// TIA Portal project "PLC_FB_Portfolio" (V14)

(* hardware
DEVICE "S71500/ET200MP station_1"  S7-1500 station
   slot 0: "Rail_0"  Rack  6ES7 590-1***0-0AA0
   slot 1: "PLC_1"  CPU 1511-1 PN  6ES7 511-1AK01-0AB0  V2.1
      slot 3: "CPU display_1"  6ES7591-1AA00-0AA0
*)

// ===== PLC "PLC_1"  CPU 1511-1 PN =====

VAR_GLOBAL   // PLC tag table "Default tag table"
   "Btn1_Start" AT %I0.0 : Bool;
   "Btn1_Stop" AT %I0.1 : Bool;
   "Btn2_Start" AT %I0.2 : Bool;
   "Btn2_Stop" AT %I0.3 : Bool;
   "BtnToggle1" AT %I0.4 : Bool;
   "BtnToggle2" AT %I0.5 : Bool;
   "FaultSim" AT %I0.6 : Bool;
   "ResetSim" AT %I0.7 : Bool;
   "Motor1" AT %Q0.0 : Bool;
   "Motor2" AT %Q0.1 : Bool;
   "Toggle1" AT %Q0.2 : Bool;
   "Toggle2" AT %Q0.3 : Bool;
END_VAR

DATA_BLOCK "FB_Toggle_DB_1"   // DB1
{ S7_Optimized_Access := 'TRUE' }
VERSION : 0.1
// stored: InstanceOfName FB_Toggle
"FB_Toggle"
BEGIN
END_DATA_BLOCK

DATA_BLOCK "FB_Toggle_DB_2"   // DB2
{ S7_Optimized_Access := 'TRUE' }
VERSION : 0.1
// stored: InstanceOfName FB_Toggle
"FB_Toggle"
BEGIN
END_DATA_BLOCK

DATA_BLOCK "FB_Motor_Latch_DB_1"   // DB3
{ S7_Optimized_Access := 'TRUE' }
VERSION : 0.1
// stored: InstanceOfName FB_Motor_Latch
"FB_Motor_Latch"
BEGIN
END_DATA_BLOCK

DATA_BLOCK "FB_Motor_Latch_DB_2"   // DB4
{ S7_Optimized_Access := 'TRUE' }
VERSION : 0.1
// stored: InstanceOfName FB_Motor_Latch
"FB_Motor_Latch"
BEGIN
END_DATA_BLOCK

FUNCTION_BLOCK "FB_Toggle"   // FB1, SCL
{ S7_Optimized_Access := 'TRUE' }
VERSION : 0.1
   VAR_INPUT
      xBtn : Bool;   // Кнопка
   END_VAR
   VAR_OUTPUT
      xOut : Bool;   // Выход
      udiToggles : UDInt;   // Счетчик переключений
   END_VAR
   VAR
      xPrevSignal : Bool;   // Память для детектера фронта
   END_VAR
BEGIN
   IF #xBtn AND NOT #xPrevSignal THEN  // фронт кнопки
       #xOut := NOT #xOut;
       #udiToggles := #udiToggles + 1;
   END_IF;

   #xPrevSignal := #xBtn;  // запоминаем для следующего вызова
END_FUNCTION_BLOCK

FUNCTION_BLOCK "FB_Motor_Latch"   // FB2, SCL
{ S7_Optimized_Access := 'TRUE' }
VERSION : 0.1
   VAR_INPUT
      xStart : Bool;   // кнопка ПУСК (фронт = команда пуска)
      xStop : Bool;   // кнопка СТОП (уровень, приоритет)
      xFault : Bool;   // авария - сброс и блокировка счета
      xReset : Bool;   // сброс счетчика пусков
   END_VAR
   VAR_OUTPUT
      xMotor : Bool;   // выход на двигатель
      xRunning : Bool;   // = xMotor AND NOT xFAult
      udiStarts : UDInt;   // счетчик успешных пусков
   END_VAR
   VAR
      xPrevStart : Bool;   // память для детектора фронта
   END_VAR
BEGIN
   // приоритет: авария > стоп > пуск
   IF #xFault OR #xStop THEN
       #xMotor := FALSE;
   ELSIF #xStart AND NOT #xPrevStart THEN  // фронт пуска
       IF NOT #xMotor THEN
           #udiStarts := #udiStarts + 1;
       END_IF;
       #xMotor := TRUE;
   END_IF;

   #xRunning := #xMotor AND NOT #xFault;

   IF #xReset THEN
       #udiStarts := 0;
   END_IF;

   #xPrevStart := #xStart;  // запоминаем для следующего вызова
END_FUNCTION_BLOCK

ORGANIZATION_BLOCK "Main"   // OB1, SCL, ProgramCycle
TITLE = "Main Program Sweep (Cycle)"
{ S7_Optimized_Access := 'TRUE' }
VERSION : 0.1
   VAR_INPUT
      Initial_Call : Bool;   // Initial call of this OB
      Remanence : Bool;   // =True, if remanent data are available
   END_VAR
BEGIN
   "FB_Toggle_DB_1"(xBtn:="BtnToggle1",
                    xOut=>"Toggle1");

   "FB_Toggle_DB_2"(xBtn:="BtnToggle2",
                    xOut=>"Toggle2");

   "FB_Motor_Latch_DB_1"(xStart:="Btn1_Start",
                         xStop:="Btn1_Stop",
                         xFault:="FaultSim",
                         xReset:="ResetSim",
                         xMotor=>"Motor1");

   "FB_Motor_Latch_DB_2"(xStart:="Btn2_Start",
                         xStop:="Btn2_Stop",
                         xFault:="FaultSim",
                         xReset:="ResetSim",
                         xMotor=>"Motor2");
END_ORGANIZATION_BLOCK